Fanuc KAREL source: KA00037.KL

PROGRAM KA00037
%NOLOCKGROUP
VAR
  SRC: STRING[80]
  DST: INTEGER
BEGIN
  SRC = 'A'
  DST = SRC
END KA00037
